Fanuc KAREL source: kc00023.KL

-- PROVISIONAL review KL for V770-1; original PC SHA256 c48601d3edb84c568939d9288448a26a09853cdc1d92399842304e9d84bc4267
-- Incomplete behavior may be omitted. Consult companion uncertainty JSON. Do not deploy.
PROGRAM KC00023
%NOLOCKGROUP
BEGIN
  -- UNRESOLVED_PC offsets 0-1; opcodes 7B
  -- UNRESOLVED_PC offsets 6-20; opcodes 2D,9D,52,2F
  -- UNRESOLVED_PC offsets 25-29; opcodes 7F
  -- UNRESOLVED_PC offsets 34-42; opcodes 3F,75
  -- UNRESOLVED_PC offsets 47-56; opcodes 3F,75
  -- UNRESOLVED_PC offsets 61-88; opcodes 27,73,73,22,24,AA,26
  -- UNRESOLVED_PC offsets 93-97; opcodes 7F
END KC00023
